(* IEC 61131-3 sources: Lasal-MCP/examples/SampleSource/5_ClassInputOutputSolution/Stations/MachineControl/MachineControl/Class/Visualize, 1 file *)

(* ---- Visualize.st ---- *)
(*!
<Class
	Name               = "Visualize"
	Revision           = "0.0"
	RealtimeTask       = "false"
	CyclicTask         = "false"
	BackgroundTask     = "false"
	Sigmatek           = "false"
	OSInterface        = "false"
	HighPriority       = "false"
	Automatic          = "false"
	UpdateMode         = "Prescan"
	SharedCommandTable = "true"
	Objectsize         = "(324,120)">
	<Channels>
		<Server Name="ClassSvr" Visualized="true" Initialize="false" WriteProtected="false" Retentive="false"/>
		<Server Name="ClientVisu" Visualized="true" Initialize="false" WriteProtected="false" Retentive="false"/>
		<Client Name="Client" Required="false" Internal="false"/>
	</Channels>
</Class>
*)
Visualize : CLASS
  //Servers:
	ClassSvr 	: SvrChCmd_DINT;
	ClientVisu 	: SvrCh_DINT;
  //Clients:
	Client 	: CltCh_DINT;
  //Variables:
  //Functions:

	FUNCTION VIRTUAL GLOBAL ClientVisu::Read
		VAR_OUTPUT
			output (EAX) 	: DINT;
		END_VAR;
  //Tables:
	FUNCTION @STD
		VAR_OUTPUT
			ret_code	: CONFSTATES;
		END_VAR;
	FUNCTION GLOBAL TAB @CT_;
END_CLASS;

FUNCTION VIRTUAL GLOBAL Visualize::ClientVisu::Read
	VAR_OUTPUT
		output (EAX) 	: DINT;
	END_VAR

	ClientVisu := Client;

	output := ClientVisu;

END_FUNCTION
